Staubli VAL3: initJogMode.pgx

public program initJogMode()
  local num l_i
begin
   for l_i = 0 to size(sShowType)-1
    sShowType[l_i]=sCartisiam[l_i]
  endFor
end
